(* IEC 61131-3 sources: SRCI_CLIENT_PLC/RobotLibrary/Library/POUs/ConveyorTracking/MC_ActivateConveyorTracking/Structures, 4 files *)

(* ---- ActivateConveyorTrackingOutCmd.st ---- *)
{attribute 'pack_mode' := '1'}
// -------------------------------------------------------------------------
//  SRCI Robot Library
// -------------------------------------------------------------------------
//
//  Object:      ActivateConveyorTrackingOutCmd
//  Author:      Thorsten Brach
//  Date:        2024-06-11
//
//  Description:
//
//
//  Copyright:
//    (C) 2024 Thorsten Brach. All rights reserved
//             Licensed under the MIT License.
//
//  Disclaimer:
//    This project is provided without any guarantee and can be used for
//    private and commercial purposes. Any use is at the user’s
//    own risk and responsibility.
//
// -------------------------------------------------------------------------
TYPE ActivateConveyorTrackingOutCmd :
STRUCT
  /// Current status of "ConveyorTracking" according to Table 6-454
  TrackingStatus     : TrackingStatus;
  /// Relates to "ConnectionMode" 1 – "RC connected": Traveled distance of assigned conveyor since ConveyorTracking has been activated (offset)
  RCEncoderValue     : REAL;
END_STRUCT
END_TYPE

(* ---- ActivateConveyorTrackingParCmd.st ---- *)
{attribute 'pack_mode' := '1'}
// -------------------------------------------------------------------------
//  SRCI Robot Library
// -------------------------------------------------------------------------
//
//  Object:      ActivateConveyorTrackingParCmd
//  Author:      Thorsten Brach
//  Date:        2024-06-11
//
//  Description:
//
//
//  Copyright:
//    (C) 2024 Thorsten Brach. All rights reserved
//             Licensed under the MIT License.
//
//  Disclaimer:
//    This project is provided without any guarantee and can be used for
//    private and commercial purposes. Any use is at the user’s
//    own risk and responsibility.
//
// -------------------------------------------------------------------------
TYPE ActivateConveyorTrackingParCmd :
STRUCT
  /// Index of assigned conveyor
  ConveyorNo         : USINT; // ST-FIX F175: ConveyorNo / ConnectionMode are USINT (6.3.26 application layer and CML; the SINT of the telegram table 6-460 is a copy error, all other conveyor telegrams have USINT)
  /// Specifies encoder connection setup (at least one option must be supported)
  ConnectionMode     : ConnectionMode;
  /// Relates to "ConnectionMode" 1 – "PLC connected": Value of the encoder connected to the conveyor belt
  PLCEncoderValue    : REAL;
END_STRUCT
END_TYPE

(* ---- ActivateConveyorTrackingRecvData.st ---- *)
{attribute 'pack_mode' := '1'}
// -------------------------------------------------------------------------
//  SRCI Robot Library
// -------------------------------------------------------------------------
//
//  Object:      ActivateConveyorTrackingRecvData
//  Author:      Thorsten Brach
//  Date:        2024-06-11
//
//  Description:
//
//
//  Copyright:
//    (C) 2024 Thorsten Brach. All rights reserved
//             Licensed under the MIT License.
//
//  Disclaimer:
//    This project is provided without any guarantee and can be used for
//    private and commercial purposes. Any use is at the user’s
//    own risk and responsibility.
//
// -------------------------------------------------------------------------
TYPE ActivateConveyorTrackingRecvData EXTENDS RspHeader :
STRUCT
  /// Maximum error of deviation of the TCP position
  /// from the fix point in world coordinate system
  /// If not supported: • -1
  TrackingStatus : TrackingStatus;
END_STRUCT
END_TYPE

(* ---- ActivateConveyorTrackingSendData.st ---- *)
{attribute 'pack_mode' := '1'}
// -------------------------------------------------------------------------
//  SRCI Robot Library
// -------------------------------------------------------------------------
//
//  Object:      ActivateConveyorTrackingSendData
//  Author:      Thorsten Brach
//  Date:        2024-06-11
//
//  Description:
//
//
//  Copyright:
//    (C) 2024 Thorsten Brach. All rights reserved
//             Licensed under the MIT License.
//
//  Disclaimer:
//    This project is provided without any guarantee and can be used for
//    private and commercial purposes. Any use is at the user’s
//    own risk and responsibility.
//
// -------------------------------------------------------------------------
TYPE ActivateConveyorTrackingSendData EXTENDS CmdHeader:
STRUCT
  /// Index of assigned conveyor
  ConveyorNo     : USINT; // ST-FIX F175: ConveyorNo / ConnectionMode are USINT (6.3.26 application layer and CML; the SINT of the telegram table 6-460 is a copy error, all other conveyor telegrams have USINT)
  /// Specifies encoder connection setup (at least one option must be supported)
  ConnectionMode : USINT; // ST-FIX F175: ConveyorNo / ConnectionMode are USINT (6.3.26 application layer and CML; the SINT of the telegram table 6-460 is a copy error, all other conveyor telegrams have USINT)
END_STRUCT
END_TYPE
